(* IEC 61131-3 sources: Lasal-MCP/examples/SampleSource/LASALScreenAdvancedSolution/LASALScreenAdvancedSolution/LASALScreenAdvacnedSolution/Stations/MachineControl/MachineControl/Network, 1 file *)

(* ---- ConfigObjects.st ---- *)
FUNCTION GLOBAL TAB TASK_CONF
_K_TASK, _K_REAL,
_K_END_VAR,

_K_TASK, _K_CYCLIC,
_K_END_VAR,

_K_TASK, _K_BACKGROUND,
_K_END_VAR,

_K_END_CONF
END_FUNCTION

FUNCTION GLOBAL TAB IPR_CONF
_K_IPR
	0$UINT,
_K_END_VAR,
_K_END_CONF
END_FUNCTION

FUNCTION GLOBAL TAB CONFIG_TABLES
00080$UINT,
0$UINT, 0, 11, "_ALARMX0PARA",
0$UINT, 0, 20, "_ALARMXBUFFER",
0$UINT, 0, 4, "_CAN",
0$UINT, 1, 10, "_CANLIB",
0$UINT, 1, 4, "_CHECKONLINESTATUS",
0$UINT, 1, 0, "_CHECKSUM",
0$UINT, 1, 20, "_FILESYS",
0$UINT, 1, 1, "_MULTITASK",
0$UINT, 0, 5, "_OSKERNEL",
0$UINT, 1, 34, "_SERLIB",
0$UINT, 1, 0, "_SIG_LSL_CMULTIMASTERSTATE",
0$UINT, 0, 0, "_STDLIB",
0$UINT, 2, 1, "_SYNCTIMEPLC",
0$UINT, 0, 9, "_SYSDATETIME",
0$UINT, 0, 0, "_SYSDATETIME2",
0$UINT, 1, 1, "_TASKOBJECTCONTROL",
0$UINT, 1, 20, "AI043",
0$UINT, 1, 40, "AM441",
0$UINT, 1, 21, "ASCII_BIN",
0$UINT, 1, 24, "BUSINTERFACESDIAS",
0$UINT, 2, 1, "BUSINTERFACESDIASINTERNAL",
0$UINT, 1, 1, "CP111_IOS",
0$UINT, 1, 1, "CP112_IOS",
0$UINT, 0, 4, "CRITICALSECTION",
0$UINT, 1, 1, "DATAMANAGER",
0$UINT, 1, 0, "DATAMANAGERFIFO",
0$UINT, 1, 0, "DATAMANAGERPRIORITY",
0$UINT, 1, 33, "DI202",
0$UINT, 2, 33, "DIASMASTER",
0$UINT, 1, 83, "DIASMASTERC",
0$UINT, 2, 25, "DIASMASTERMAIN",
0$UINT, 1, 0, "DIASMASTERPOSTSCAN",
0$UINT, 1, 14, "DM161",
0$UINT, 1, 11, "EEPROM",
0$UINT, 1, 2, "GETOSVERSION",
0$UINT, 0, 2, "GETTASKHANDLE",
0$UINT, 1, 21, "HUB_BASE",
0$UINT, 2, 11, "HUB_BASE_ROOT",
0$UINT, 2, 36, "HWBASE",
0$UINT, 2, 56, "HWBASECDIAS",
0$UINT, 1, 0, "HWCLOGGING",
0$UINT, 5, 19, "HWCONTROL",
0$UINT, 1, 10, "HWCONTROLBASE",
0$UINT, 1, 0, "HWRTPOSTSCAN",
0$UINT, 1, 6, "I2CCDIAS",
0$UINT, 1, 22, "MERKEREX",
0$UINT, 1, 75, "PLC_INFO",
0$UINT, 1, 3, "RAM",
0$UINT, 1, 9, "RAMFILE",
0$UINT, 1, 1, "RAMRINGBUFFER",
0$UINT, 1, 22, "SAFETYBASEFSOE",
0$UINT, 3, 19, "SAFETYCDIAS_BASE",
0$UINT, 2, 24, "SAFETYMANAGER",
0$UINT, 1, 4, "SAFETYUDP",
0$UINT, 1, 36, "SCP111",
0$UINT, 1, 60, "SDIASBASE",
0$UINT, 1, 10, "SDIASHUBBASE",
0$UINT, 1, 97, "SDIASMANAGER",
0$UINT, 2, 6, "SDIASPLC",
0$UINT, 1, 9, "SDIASSAFETYBASE",
0$UINT, 1, 25, "SDIASSAFETYMANAGERFSOE",
0$UINT, 1, 11, "SDM081",
0$UINT, 0, 37, "SIGCLIB",
0$UINT, 1, 11, "STRING",
0$UINT, 1, 85, "STRINGINTERNAL",
0$UINT, 1, 21, "SYNCCALL",
0$UINT, 0, 1, "SYSTEM",
0$UINT, 0, 0, "TANK",
0$UINT, 1, 17, "TCPCOMMUNICATION",
0$UINT, 1, 0, "TCPCOMMUNICATIONLOGFILTER",
0$UINT, 1, 44, "TO127",
0$UINT, 1, 1, "USERALARMGENERATOR",
0$UINT, 2, 18, "VARAN_BASE",
0$UINT, 3, 4, "VARANMANAGER",
0$UINT, 2, 4, "VARANMANAGER_1",
0$UINT, 2, 6, "VARANMANAGER_2",
0$UINT, 1, 25, "VARANMANAGER_BASE",
0$UINT, 1, 3, "VIRTUALBASEINIT",
0$UINT, 2, 11, "WATCHDOGDIAS",
0$UINT, 1, 1, "XXXBASE_IOS",
ONE_CFG$UINT, 0, 0, "ONE_HW_Network",
ONE_CFG$UINT, 1, 0, "ONE_STDAlarm",
ONE_CFG$UINT, 1, 0, "ONE_STDCommunicationToHMI",
ONE_CFG$UINT, 1, 0, "ONE_STDPLCInfoPLC",
ONE_CFG$UINT, 2, 0, "ONE_STDTimeSync",
ONE_CFG$UINT, 0, 0, "ONE_TankNet",
TASK_CFG$UINT, 0, 0, "TASK_CONF",
IPR_CFG$UINT, 0, 0, "IPR_CONF",
PRJ_CFG$UINT, 0, 0, "MachineControl",
END_FUNCTION

#ifdef __LSLLDR_IOELEMENTS__
FUNCTION GLOBAL TAB _IO_ELEMENTS_TAB
0001$UINT, 0001$UINT,
"Potentiometer", "AI0431.AI2",
0001$UINT,
"Potentiometer", "Tank1.ActFillLevel",
END_FUNCTION
#endif //__LSLLDR_IOELEMENTS__

FUNCTION GLOBAL TAB CH_REDIRECT_EMB_TAB
0000$UINT,
00024$UINT,
"AI043;SERIALNO", "\SERIALNOSTR.DATA",
"AM441;SERIALNO", "\SERIALNOSTR.DATA",
"BUSINTERFACESDIAS;SERIALNO", "\SERIALNOSTR.DATA",
"DI202;SERIALNO", "\SERIALNOSTR.DATA",
"DM161;SERIALNO", "\SERIALNOSTR.DATA",
"HWBASECDIAS;SERIALNO", "\SERIALNOSTR.DATA",
"PLC_INFO;APPLICATIONNAME", "\APPLINAME.DATA",
"PLC_INFO;CPUBOARDNAME", "\CPUBOARD.DATA",
"PLC_INFO;CPU_NAME", "\STRING1.DATA",
"PLC_INFO;DISPLAYNAME", "\CHASSISTYPE.DATA",
"PLC_INFO;SERNUM", "\STRING0.DATA",
"PLC_INFO;SYSINFOSTRING", "\SYSINFO.DATA",
"SAFETYCDIAS_BASE;SERIALNO", "\SERIALNOSTR.DATA",
"SCP111;DESIGNERPRJNAME", "\SDIASSAFETYMANAGERFSOE1\PROJECTNAMESTR.DATA",
"SCP111;DESIGNERPRJREV", "\SDIASSAFETYMANAGERFSOE1\PROJECTREVISIONSTR.DATA",
"SCP111;SERIALNO", "\SERIALNOSTR.DATA",
"SDIASBASE;SERIALNO", "\SERIALNOSTR.DATA",
"SDIASSAFETYBASE;SERIALNO", "\SERIALNOSTR.DATA",
"SDIASSAFETYMANAGERFSOE;DESIGNERPRJNAME", "\PROJECTNAMESTR.DATA",
"SDIASSAFETYMANAGERFSOE;DESIGNERPRJREV", "\PROJECTREVISIONSTR.DATA",
"SDM081;SERIALNO", "\SERIALNOSTR.DATA",
"TCPCOMMUNICATION;TASKNAME", "\THREADNAME.DATA",
"TO127;SERIALNO", "\SERIALNOSTR.DATA",
"VARAN_BASE;SERIALNO", "\SERIALNOSTR.DATA",
END_FUNCTION
